(* IEC 61131-3 sources: kns-pump-station/src/POUs/Field/Owen/F_Mx210AiToMa, 2 files *)

(* ---- F_Mx210AiToMa.decl.st ---- *)
// Назначение: аналоговый вход модуля ОВЕН Mx210 (МВ210-101) по Modbus → ток для PL.FB_AnalogInput.
//             «Значение (float) на входе» — FLOAT32 в двух регистрах, младшее слово первым (так их собирает
//             пример ОВЕН Example_CodesysModbusTcpMasterMx210_3517v1). Для датчика 4–20 мА модуль даёт
//             0…100 % → 4…20 мА. Старший байт 16#F0…16#FF — код ошибки входа (обрыв, КЗ, нет данных; РЭ
//             МВ210-101) — NaN, как и при потере связи с модулем (решает вызывающий). Сборка targets/plc210.
// Автор:      kr0nsch
// Версия:     0.1.0
// Документ:   docs/DESIGN.md, раздел 8.4; targets/plc210/README.md
FUNCTION F_Mx210AiToMa : REAL
VAR_INPUT
    wLo : WORD;     // первый регистр (младшее слово FLOAT32)
    wHi : WORD;     // второй регистр (старшее слово; старший байт — код ошибки)
END_VAR
VAR
    uBits : PL.U_RealBits;  // NaN из битов
END_VAR

(* ---- F_Mx210AiToMa.impl.st ---- *)
IF SHR(wHi, GVL_Const.MB_BYTE_BITS) >= GVL_Const.MX210_AI_ERR_MIN THEN
    uBits.dwValue := GVL_Const.REAL_QNAN_BITS;
    F_Mx210AiToMa := uBits.rValue;
ELSE
    F_Mx210AiToMa := PL.GVL_Const.MA_ZERO
                     + F_WordsToReal(wHi := wHi, wLo := wLo) * PL.GVL_Const.MA_SPAN / PL.GVL_Const.PCT_FULL;
END_IF
